(* IEC 61131-3 sources: 2026_Projet_YGO_ExcavatriceDragage/CODE/MAIN (part 2) *)

(* ---- PRG_09_Supervision.st ---- *)
(* ═══════════════════════════════════════════════════════════════
   🖥️ PRG_09_Supervision — Échanges IHM, Stubs et Initialisation Boot
   ───────────────────────────────────────────────────────────────
   ⚙️ Exécuté par la tâche PLC en position 9.
   ✅ Regroupe tout le mapping bidirectionnel GVL_IHM / GVL_PERSISTENT.
   ✅ Expose FaultMachineReset_IHM pour tous les programmes du domaine sécurité/métier.
   🔧 REX 2026-07-07 : séparation des resets — l'ancien MachineReset_IHM (unique, câblé sur
      TOUT y compris FB_Modes/FB_Cycle) est retiré. FaultMachineReset_IHM ne couvre plus que le
      domaine sécurité/métier (Winch, Safety, Encodeurs, Benne, Joystick, Translation) ;
      FB_Modes/FB_Cycle ont chacun leur propre Reset dédié (GVL_IHM.Modes.ModeReset côté
      PRG_04_Modes, CmdResetCycle_IHM côté PRG_05_Cycle) — jamais mélangés.
   ═══════════════════════════════════════════════════════════════ *)

PROGRAM PRG_09_Supervision
VAR_OUTPUT
    FaultMachineReset_IHM : BOOL; // 🔔 Acquittement défauts domaine sécurité/métier (OR des boutons HMI) — jamais Modes/Cycle
END_VAR
VAR
    instBlink1Hz : BLINK; // 🧩 Réutilisation lib Util (Partie3 §0) — horloge clignotement système
END_VAR

// === IMPLEMENTATION (corps du PROGRAM PRG_09_Supervision) ===

// ── 0. HORLOGE CLIGNOTEMENT SYSTÈME (GVL_Global.BlinkClock) ───────────────
// 🧩 Réutilisation lib Util (Partie3 §0) : bloc standard BLINK, pas de TON maison —
// gère nativement un rythme allumé/éteint ASYMÉTRIQUE (TimeHigh ≠ TimeLow), contrairement
// au motif TON manuel de FB_Output.st (symétrique 500/500, propre à l'option relais).
// 🔧 REX 2026-07-16 : durées réglables sans recompiler (GVL_PERSISTENT._BlinkTimeOn/_BlinkTimeOff,
// défaut 1s allumé / 800ms éteint) — un seul rythme partagé pour tous les voyants IHM/diag qui
// clignotent pareil.
// 💡 Un voyant a besoin d'un AUTRE rythme ? Instancier son propre BLINK localement (Util) avec
// ses propres TimeHigh/TimeLow — ne pas détourner ce bit partagé pour un rythme différent.
instBlink1Hz(
    ENABLE   := TRUE,
    TIMEHIGH := _BlinkTimeOn,
    TIMELOW  := _BlinkTimeOff
);
GVL_Global.BlinkClock := instBlink1Hz.OUT;

// ── 1. ACQUISITION DES DEMANDES / BOUTONS DE L'IHM ────────────────────────
GVL_Modes_Stub.ModeRequest_IHM         := GVL_IHM.Modes.ModeRequest;
GVL_Modes_Stub.SyncEnableRequest_IHM   := GVL_IHM.Sync.SyncEnableRequest; // 🔧 REX 2026-07-08 : renommé, polarité inversée
StubTranslationPositionSelect_IHM          := GVL_IHM.TranslationM3.SelectedTargetNum;

// Signal d'acquittement défauts domaine sécurité/métier — JAMAIS Modes/Cycle (REX 2026-07-07)
FaultMachineReset_IHM := GVL_IHM.Modes.FaultMachineReset
                    OR GVL_IHM.M1TreuilRetenue.CmdReset
                    OR GVL_IHM.M2TreuilBucket.CmdReset
                    OR GVL_IHM.Bucket.CmdReset;

// 🔴 REX 2026-07-07 : au moins un défaut actif dans le domaine couvert par FaultMachineReset_IHM
// (même périmètre exact que les 17 blocs alimentés par ce reset — voir bandeau en tête de fichier).
// Sert à savoir, côté IHM, quand un appui sur FaultMachineReset est utile/attendu.
GVL_IHM.Modes.AnyFaultActive :=
       PRG_01_Diagnostics.instDiagCanOpen.Error
    OR PRG_01_Diagnostics.instDiagEthercat.Error
    OR PRG_01_Diagnostics.FB_Joystick_0.Error
    OR (NOT PRG_04_Modes.instModes.InhibitM1 AND (
           PRG_02_Encoders.instEncoderAbsM1.Error
        OR PRG_02_Encoders.instHomingM1.Error
        OR PRG_02_Encoders.instEncoderSafetyM1.Error
        OR PRG_03_Safety.instSafetyWinchM1.Error
        OR PRG_06_WinchControl.instWinchM1.Error
    ))
    OR (NOT PRG_04_Modes.instModes.InhibitM2 AND (
           PRG_02_Encoders.instEncoderAbsM2.Error
        OR PRG_02_Encoders.instHomingM2.Error
        OR PRG_02_Encoders.instEncoderSafetyM2.Error
        OR PRG_03_Safety.instSafetyWinchM2.Error
        OR PRG_06_WinchControl.instWinchM2.Error
    ))
    OR PRG_03_Safety.instSafetyTranslationM3.Error
    OR PRG_06_WinchControl.instWinchSync.Error
    OR PRG_06_WinchControl.instBucket.Error
    OR PRG_07_TranslationControl.instTranslationM3.Error
    OR PRG_10_Outputs.RedundancyTestFailed
    OR PRG_10_Outputs.EmergencyArmingFailed;

// 🧨 REX 2026-07-07 : remontée IHM de la coupure puissance amont — polarité "alarme" (TRUE=
// problème), PAS celle de PowerCutOff_A_RQ (qui est en fail-safe maintenu, TRUE=OK depuis
// l'inversion de polarité). On relit directement les .PowerCutOff sources, pas la sortie physique.
GVL_IHM.Modes.PowerCutOffActive := PRG_03_Safety.instSafetyWinchM1.PowerCutOff
                                 OR PRG_03_Safety.instSafetyWinchM2.PowerCutOff
                                 OR PRG_03_Safety.instSafetyTranslationM3.PowerCutOff
                                 OR GVL_IHM.Modes.CmdEmergencyCutOff;

// 🆕 REX 2026-07-08 : thermique frein commun M1/M2/M3 — signal UNIQUE (1 seul fil, pas de sens à
// le dupliquer par axe), remonté une seule fois au niveau global GVL_IHM (même principe que
// TopPositionSensorActive ci-dessus, PAS dans WinchM1/WinchM2/Translation).
GVL_IHM.Commun.BrakeThermalFault := NOT PRG_00_Inputs.BrakeThermalFeedback;
GVL_IHM.Commun.PhaseRotationFault := NOT PRG_00_Inputs.PhaseRotationOk; // 🆕 REX 2026-07-08 — commun M1/M2/M3, invisible IHM avant

// 🔧 REX 2026-07-07 — Séquence réarmement AU (voir DOC/AF_Partie1 v1.5 §Sécurité électrique)
// EmergencyArmingBusy couvre TOUTE la séquence (auto-test A/B + pulse + confirmation + verrouillage),
// pas seulement le pulse — ArmingSeqStep<>0 englobe déjà tout sauf le verrouillage final.
GVL_IHM.Modes.EmergencyChainOk    := PRG_00_Inputs.EmergencyChain;
GVL_IHM.Modes.PowerContactorOk    := PRG_00_Inputs.EmergencyStopOk;
GVL_IHM.Modes.EmergencyArmingBusy := (PRG_10_Outputs.ArmingSeqStep <> 0) OR PRG_10_Outputs.EmergencyArmingLockoutActive;
GVL_IHM.Modes.EmergencyArmable    := PRG_00_Inputs.EmergencyChain
                                    AND (PRG_10_Outputs.ArmingSeqStep = 0)
                                    AND NOT PRG_10_Outputs.EmergencyArmingLockoutActive
                                    AND NOT PRG_10_Outputs.RedundancyTestFailed;
GVL_IHM.Modes.RedundancyTestFailed := PRG_10_Outputs.RedundancyTestFailed;
GVL_IHM.Modes.EmergencyArmingFailed := PRG_10_Outputs.EmergencyArmingFailed;

// 🔧 REX 2026-07-07 : ancien pont IF/ELSIF vers GVL_Encoder_Stub supprimé (bugué — ne pouvait
// homer qu'un seul treuil à la fois). GVL_IHM.M1TreuilRetenue/M2.CmdHome sont désormais câblés
// directement dans PRG_02_Encoders.st (instHomingM1/M2.Home) — homing simultané possible.

// ℹ️ Calibrate joystick : lu directement depuis GVL_IHM.JoystickJOY1.Calibrate dans PRG_01_Diagnostics (ligne 48)
// PRG_01_Diagnostics.FB_Joystick_0.Calibrate := GVL_IHM.JoystickJOY1.Calibrate;  // ❌ supprimé : VAR locale non accessible en écriture (C0037)

// ── 2. INITIALISATION IHM DEPUIS GVL_PERSISTENT (Boot) ───────────────────
IF GVL_IHM.M1TreuilRetenue.TopSensorPositionM = 0.0 THEN
    GVL_IHM.M1TreuilRetenue.TopSensorPositionM  := _HomingTargetM1_M;
    GVL_IHM.M1TreuilRetenue.MaxStepDescente     := _WinchMaxStepDescent; // 🔧 REX 2026-07-08 : commun M1/M2
    GVL_IHM.M1TreuilRetenue.RampAccelRate       := _WinchM1RampAccelRate_Pct;
    GVL_IHM.M1TreuilRetenue.RampDecelNormalRate := _WinchM1RampDecelNormal_Pct;
    GVL_IHM.M1TreuilRetenue.RampDecelFastRate   := _WinchM1RampDecelFast_Pct;
    GVL_IHM.M1TreuilRetenue.CableLimitDescentM  := _CableLimitM1Descent_M;
    GVL_IHM.M1TreuilRetenue.CableLimitAscentM   := _CableLimitM1Ascent_M; // 🆕 REX 2026-07-15 (6)
    GVL_IHM.M1TreuilRetenue.SlowdownDistanceM   := _WinchSlowdownDistance_M;
    GVL_IHM.M1TreuilRetenue.SlowSpeedPct        := _WinchSlowSpeed_Pct;
END_IF;

IF GVL_IHM.M2TreuilBucket.TopSensorPositionM = 0.0 THEN
    GVL_IHM.M2TreuilBucket.TopSensorPositionM  := _HomingTargetM2_M;
    GVL_IHM.M2TreuilBucket.MaxStepDescente     := _WinchMaxStepDescent; // 🔧 REX 2026-07-08 : commun M1/M2
    GVL_IHM.M2TreuilBucket.RampAccelRate       := _WinchM2RampAccelRate_Pct;
    GVL_IHM.M2TreuilBucket.RampDecelNormalRate := _WinchM2RampDecelNormal_Pct;
    GVL_IHM.M2TreuilBucket.RampDecelFastRate   := _WinchM2RampDecelFast_Pct;
    GVL_IHM.M2TreuilBucket.CableLimitDescentM  := _CableLimitM2Descent_M;
    GVL_IHM.M2TreuilBucket.CableLimitAscentM   := _CableLimitM2Ascent_M; // 🆕 REX 2026-07-15 (6)
    GVL_IHM.M2TreuilBucket.SlowdownDistanceM   := _WinchSlowdownDistance_M;
    GVL_IHM.M2TreuilBucket.SlowSpeedPct        := _WinchSlowSpeed_Pct;
END_IF;

IF GVL_IHM.Sync.SyncToleranceM = 0.0 THEN
    GVL_IHM.Sync.SyncToleranceM         := _WinchSyncTolerance_M;
END_IF;

IF GVL_IHM.Bucket.Config.OffsetOpenM = 0.0 AND GVL_IHM.Bucket.Config.OffsetCloseM = 0.0 THEN
    GVL_IHM.Bucket.Config := _BucketConfig;
    GVL_IHM.Bucket.TimeoutDuration := T#30s;
END_IF;

IF GVL_IHM.Commun.LimitLegalDepthMinAllowed = 0.0 THEN
    GVL_IHM.Commun.LimitLegalDepthMinAllowed := _LimitLegalDepthMinAllowed_M;
    GVL_IHM.Commun.LimitLegalEnabled         := _LimitLegalEnabled;
END_IF;

// 🆕 REX 2026-07-15 (10) — BUG CORRIGÉ (retour terrain) : WinchMaxStepFwd/Rev (essais progressifs
// IHM_MANU, TEMPORAIRE) n'avaient jamais de boot-init, contrairement à tous les autres réglages
// IHM ci-dessus — restaient à 0 (défaut INT) en permanence. Le bornage de PRG_06_WinchControl
// traitait ce 0 comme "invalide" et le remplaçait SILENCIEUSEMENT par 5 (aucune restriction),
// sans jamais corriger l'affichage IHM : l'opérateur voyait "0" (lu comme restrictif) alors que
// la vitesse réellement appliquée était pleine échelle — d'où les contacteurs qui commutaient
// normalement malgré un "0" à l'écran. GVL_IHM.IHM_MANU est déjà RETAIN (ST_IHM_MANU) — pas besoin
// de miroir GVL_PERSISTENT (dérogation temporaire, pas un réglage machine permanent, voir
// IHM_MANU_Journal_Modifications.md §10).
IF GVL_IHM.IHM_MANU.WinchMaxStepFwd = 0 THEN
    GVL_IHM.IHM_MANU.WinchMaxStepFwd := 5;
END_IF;
IF GVL_IHM.IHM_MANU.WinchMaxStepRev = 0 THEN
    GVL_IHM.IHM_MANU.WinchMaxStepRev := 2;
END_IF;

IF GVL_IHM.Modes.ModeRequest = E_Mode.DISABLE THEN
    GVL_IHM.Modes.ModeRequest := E_Mode.MAINT_N1;
END_IF;

// ── 3. PROPAGATION DES RÉGLAGES IHM → PERSISTANCE ───────────────────────
_HomingTargetM1_M           := GVL_IHM.M1TreuilRetenue.TopSensorPositionM;
_HomingTargetM2_M           := GVL_IHM.M2TreuilBucket.TopSensorPositionM;
// 🔧 REX 2026-07-08 : MaxStepDescente désormais commun M1/M2 — voir bloc miroir bidirectionnel
// ci-dessous (même pattern que CableLimitDescentM/SlowdownDistanceM/SlowSpeedPct), plus de
// propagation à sens unique séparée par treuil ici.
_WinchM1RampAccelRate_Pct   := GVL_IHM.M1TreuilRetenue.RampAccelRate;
_WinchM1RampDecelNormal_Pct := GVL_IHM.M1TreuilRetenue.RampDecelNormalRate;
_WinchM1RampDecelFast_Pct   := GVL_IHM.M1TreuilRetenue.RampDecelFastRate;
_WinchM2RampAccelRate_Pct   := GVL_IHM.M2TreuilBucket.RampAccelRate;
_WinchM2RampDecelNormal_Pct := GVL_IHM.M2TreuilBucket.RampDecelNormalRate;
_WinchM2RampDecelFast_Pct   := GVL_IHM.M2TreuilBucket.RampDecelFastRate;
// ⚠️ REX 2026-07-08 (5) — PIÈGE pont IHM→PERSISTENT découvert lors de l'audit : cette ligne
// écrase _WinchSyncTolerance_M avec GVL_IHM.Sync.SyncToleranceM À CHAQUE SCAN.
// Si on change UNIQUEMENT la valeur par défaut dans GVL_PERSISTENT.st (ou ST_SyncHMI.st), ça ne
// suffit pas : la valeur restaurée au boot (bloc §2 ci-dessus, `IF ... = 0.0 THEN`) ne s'applique
// que si le RETAIN IHM est à 0.0 (premier démarrage) — sinon l'ancienne valeur IHM re-propage ici
// et écrase silencieusement toute nouvelle valeur par défaut au scan suivant.
_WinchSyncTolerance_M       := GVL_IHM.Sync.SyncToleranceM;
_BucketConfig              := GVL_IHM.Bucket.Config;

// 🔧 REX 2026-07-08 (demande utilisateur) : MaxStepDescente commun M1/M2 — même profil de
// déplacement des 2 treuils, même pattern miroir que CableLimitDescentM ci-dessous.
IF GVL_IHM.M1TreuilRetenue.MaxStepDescente <> _WinchMaxStepDescent THEN
    _WinchMaxStepDescent := GVL_IHM.M1TreuilRetenue.MaxStepDescente;
ELSIF GVL_IHM.M2TreuilBucket.MaxStepDescente <> _WinchMaxStepDescent THEN
    _WinchMaxStepDescent := GVL_IHM.M2TreuilBucket.MaxStepDescente;
END_IF;
GVL_IHM.M1TreuilRetenue.MaxStepDescente := _WinchMaxStepDescent;
GVL_IHM.M2TreuilBucket.MaxStepDescente := _WinchMaxStepDescent;

IF GVL_IHM.M1TreuilRetenue.CableLimitDescentM <> _CableLimitM1Descent_M THEN
    _CableLimitM1Descent_M := GVL_IHM.M1TreuilRetenue.CableLimitDescentM;
END_IF;
GVL_IHM.M1TreuilRetenue.CableLimitDescentM := _CableLimitM1Descent_M;

IF GVL_IHM.M2TreuilBucket.CableLimitDescentM <> _CableLimitM2Descent_M THEN
    _CableLimitM2Descent_M := GVL_IHM.M2TreuilBucket.CableLimitDescentM;
END_IF;
GVL_IHM.M2TreuilBucket.CableLimitDescentM := _CableLimitM2Descent_M;

// 🆕 REX 2026-07-15 (6) — même pattern miroir bidirectionnel que CableLimitDescentM ci-dessus.
IF GVL_IHM.M1TreuilRetenue.CableLimitAscentM <> _CableLimitM1Ascent_M THEN
    _CableLimitM1Ascent_M := GVL_IHM.M1TreuilRetenue.CableLimitAscentM;
END_IF;
GVL_IHM.M1TreuilRetenue.CableLimitAscentM := _CableLimitM1Ascent_M;

IF GVL_IHM.M2TreuilBucket.CableLimitAscentM <> _CableLimitM2Ascent_M THEN
    _CableLimitM2Ascent_M := GVL_IHM.M2TreuilBucket.CableLimitAscentM;
END_IF;
GVL_IHM.M2TreuilBucket.CableLimitAscentM := _CableLimitM2Ascent_M;

IF GVL_IHM.M1TreuilRetenue.SlowdownDistanceM <> _WinchSlowdownDistance_M THEN
    _WinchSlowdownDistance_M := GVL_IHM.M1TreuilRetenue.SlowdownDistanceM;
ELSIF GVL_IHM.M2TreuilBucket.SlowdownDistanceM <> _WinchSlowdownDistance_M THEN
    _WinchSlowdownDistance_M := GVL_IHM.M2TreuilBucket.SlowdownDistanceM;
END_IF;
GVL_IHM.M1TreuilRetenue.SlowdownDistanceM := _WinchSlowdownDistance_M;
GVL_IHM.M2TreuilBucket.SlowdownDistanceM := _WinchSlowdownDistance_M;

IF GVL_IHM.M1TreuilRetenue.SlowSpeedPct <> _WinchSlowSpeed_Pct THEN
    _WinchSlowSpeed_Pct := GVL_IHM.M1TreuilRetenue.SlowSpeedPct;
ELSIF GVL_IHM.M2TreuilBucket.SlowSpeedPct <> _WinchSlowSpeed_Pct THEN
    _WinchSlowSpeed_Pct := GVL_IHM.M2TreuilBucket.SlowSpeedPct;
END_IF;
GVL_IHM.M1TreuilRetenue.SlowSpeedPct := _WinchSlowSpeed_Pct;
GVL_IHM.M2TreuilBucket.SlowSpeedPct := _WinchSlowSpeed_Pct;

_LimitLegalDepthMinAllowed_M := GVL_IHM.Commun.LimitLegalDepthMinAllowed;
_LimitLegalEnabled         := GVL_IHM.Commun.LimitLegalEnabled;
// 🔧 REX 2026-07-07 : plus de garde Mode=SEMI_AUTO, cohérent avec PRG_06_WinchControl.st §5
// (la limite légale s'applique désormais dans tous les modes dès qu'elle est activée).
GVL_IHM.Commun.LimitLegalReached         := _LimitLegalEnabled
                                            AND ((NOT PRG_04_Modes.instModes.InhibitM1 AND (PRG_02_Encoders.instEncoderScaleM1.CablePosM <= _LimitLegalDepthMinAllowed_M))
                                                 OR (NOT PRG_04_Modes.instModes.InhibitM2 AND (PRG_02_Encoders.instEncoderScaleM2.CablePosM <= _LimitLegalDepthMinAllowed_M)));

GVL_IHM.Commun.TopPositionSensorActive   := NOT PRG_00_Inputs.TopPositionSensor;

// ── 4. BYPASS DE SIMULATION POUR L'IHM (état effectif par device, voir AF_Partie13) ──────
GVL_IHM.M1TreuilRetenue.BypassContactorFeedback := GVL_Simulation.SimulationModeActive AND NOT GVL_Simulation.ContactorFeedbackM1_IsReal;
GVL_IHM.M2TreuilBucket.BypassContactorFeedback := GVL_Simulation.SimulationModeActive AND NOT GVL_Simulation.ContactorFeedbackM2_IsReal;
GVL_IHM.TranslationM3.BypassContactorFeedback := GVL_Simulation.SimulationModeActive AND NOT GVL_Simulation.ContactorFeedbackM3_IsReal;
GVL_IHM.M1TreuilRetenue.BypassSlackCable        := GVL_Simulation.SimulationModeActive AND NOT GVL_Simulation.SlackCableSwitch_IsReal;
GVL_IHM.M2TreuilBucket.BypassSlackCable        := GVL_Simulation.SimulationModeActive AND NOT GVL_Simulation.SlackCableSwitch_IsReal;
GVL_IHM.M1TreuilRetenue.BypassTopPositionSensor := GVL_Simulation.SimulationModeActive AND NOT GVL_Simulation.TopPositionSensor_IsReal;
GVL_IHM.M2TreuilBucket.BypassTopPositionSensor := GVL_Simulation.SimulationModeActive AND NOT GVL_Simulation.TopPositionSensor_IsReal;

// ── 5. MAPPING ÉTATS TREUIL M1 → IHM ─────────────────────────────────────
GVL_IHM.M1TreuilRetenue.PositionM                := PRG_02_Encoders.instEncoderScaleM1.CablePosM;
GVL_IHM.M1TreuilRetenue.SpeedRefPct              := PRG_06_WinchControl.instWinchM1.SpeedRamp.Current;
GVL_IHM.M1TreuilRetenue.StepNumber               := PRG_06_WinchControl.instWinchM1.StepNumber;
GVL_IHM.M1TreuilRetenue.FBState                  := PRG_06_WinchControl.instWinchM1.State;
GVL_IHM.M1TreuilRetenue.Ready                    := PRG_06_WinchControl.instWinchM1.Ready;
GVL_IHM.M1TreuilRetenue.Busy                     := PRG_06_WinchControl.instWinchM1.Busy;
GVL_IHM.M1TreuilRetenue.Done                     := PRG_06_WinchControl.instWinchM1.Done;
GVL_IHM.M1TreuilRetenue.Error                    := PRG_06_WinchControl.instWinchM1.Error;
GVL_IHM.M1TreuilRetenue.ErrorId                  := PRG_06_WinchControl.instWinchM1.ErrorId;
GVL_IHM.M1TreuilRetenue.RelayFwd                 := PRG_06_WinchControl.instWinchM1.RelayFwd;
GVL_IHM.M1TreuilRetenue.RelayRev                 := PRG_06_WinchControl.instWinchM1.RelayRev;
GVL_IHM.M1TreuilRetenue.Contactor1               := PRG_06_WinchControl.instWinchM1.Contactor1;
GVL_IHM.M1TreuilRetenue.Contactor2               := PRG_06_WinchControl.instWinchM1.Contactor2;
GVL_IHM.M1TreuilRetenue.Contactor3               := PRG_06_WinchControl.instWinchM1.Contactor3;
GVL_IHM.M1TreuilRetenue.Contactor4               := PRG_06_WinchControl.instWinchM1.Contactor4;
GVL_IHM.M1TreuilRetenue.BrakeCmd                 := PRG_06_WinchControl.instWinchM1.BrakeCmd;
GVL_IHM.M1TreuilRetenue.Homed                    := PRG_02_Encoders.instHomingM1.Homed;
GVL_IHM.M1TreuilRetenue.SafeStopActive           := PRG_03_Safety.instSafetyWinchM1.SafeStop;
GVL_IHM.M1TreuilRetenue.ForbidDescentActive      := PRG_06_WinchControl.ForbidDescentM1_Active;
GVL_IHM.M1TreuilRetenue.ForbidAscentActive       := PRG_03_Safety.instSafetyWinchM1.ForbidAscent;
GVL_IHM.M1TreuilRetenue.SlackCableDetected       := NOT PRG_00_Inputs.SlackCableSwitch;
GVL_IHM.M1TreuilRetenue.ThermalFault             := NOT PRG_00_Inputs.M1ThermalFeedback;
GVL_IHM.M1TreuilRetenue.EncoderFault             := NOT PRG_02_Encoders.instEncoderAbsM1.EncoderAvailable OR PRG_02_Encoders.instEncoderSafetyM1.EncoderIncoherent;
GVL_IHM.M1TreuilRetenue.CableLimitDescentReached := (PRG_03_Safety.instSafetyWinchM1.ErrorId AND 16#0040) <> 16#0000;
GVL_IHM.M1TreuilRetenue.CableLimitAscentReached  := PRG_06_WinchControl.CableLimitAscentM1Reached; // 🆕 REX 2026-07-15 (8)
GVL_IHM.M1TreuilRetenue.ContactorsCheck          := PRG_06_WinchControl.instWinchM1.ContactorsCheck; // 🔧 REX 2026-07-07
GVL_IHM.M1TreuilRetenue.BrakeContactorCheck      := PRG_06_WinchControl.instWinchM1.BrakeContactorCheck;

GVL_IHM.M1TreuilRetenue.Encoder.RawPos           := PRG_02_Encoders.instEncoderAbsM1.RawPos;
GVL_IHM.M1TreuilRetenue.Encoder.Alarms           := PRG_02_Encoders.instEncoderAbsM1.AlarmsIn;
GVL_IHM.M1TreuilRetenue.Encoder.Warnings         := PRG_02_Encoders.instEncoderAbsM1.WarningsIn;
GVL_IHM.M1TreuilRetenue.Encoder.SlaveOperational := PRG_02_Encoders.instEncoderAbsM1.SlaveOperational;
GVL_IHM.M1TreuilRetenue.Encoder.PresetTriggerCmd := PRG_02_Encoders.instEncoderAbsM1.PresetTriggerCmd;
GVL_IHM.M1TreuilRetenue.Encoder.PresetValueOut   := PRG_02_Encoders.instEncoderAbsM1.PresetValueOut;
GVL_IHM.M1TreuilRetenue.Encoder.Error            := PRG_02_Encoders.instEncoderAbsM1.Error;
GVL_IHM.M1TreuilRetenue.Encoder.ErrorId          := PRG_02_Encoders.instEncoderAbsM1.ErrorId;
GVL_IHM.M1TreuilRetenue.SafetyError              := PRG_03_Safety.instSafetyWinchM1.Error;
GVL_IHM.M1TreuilRetenue.SafetyErrorId            := PRG_03_Safety.instSafetyWinchM1.ErrorId;
GVL_IHM.M1TreuilRetenue.MecaADriftM              := PRG_03_Safety.instSafetyWinchM1.MecaADriftM;      // 🆕 REX 2026-07-08
GVL_IHM.M1TreuilRetenue.MecaCDriftM              := PRG_03_Safety.instSafetyWinchM1.MecaCDriftM;      // 🆕 REX 2026-07-08
GVL_IHM.M1TreuilRetenue.MecaBElapsedTime         := PRG_03_Safety.instSafetyWinchM1.MecaBElapsedTime; // 🆕 REX 2026-07-08
GVL_IHM.M1TreuilRetenue.InhibitActive            := PRG_04_Modes.instModes.InhibitM1; // 🆕 REX 2026-07-08

// ── 6. MAPPING ÉTATS TREUIL M2 → IHM ─────────────────────────────────────
GVL_IHM.M2TreuilBucket.PositionM                := PRG_02_Encoders.instEncoderScaleM2.CablePosM;
GVL_IHM.M2TreuilBucket.SpeedRefPct              := PRG_06_WinchControl.instWinchM2.SpeedRamp.Current;
GVL_IHM.M2TreuilBucket.StepNumber               := PRG_06_WinchControl.instWinchM2.StepNumber;
GVL_IHM.M2TreuilBucket.FBState                  := PRG_06_WinchControl.instWinchM2.State;
GVL_IHM.M2TreuilBucket.Ready                    := PRG_06_WinchControl.instWinchM2.Ready;
GVL_IHM.M2TreuilBucket.Busy                     := PRG_06_WinchControl.instWinchM2.Busy;
GVL_IHM.M2TreuilBucket.Done                     := PRG_06_WinchControl.instWinchM2.Done;
GVL_IHM.M2TreuilBucket.Error                    := PRG_06_WinchControl.instWinchM2.Error;
GVL_IHM.M2TreuilBucket.ErrorId                  := PRG_06_WinchControl.instWinchM2.ErrorId;
GVL_IHM.M2TreuilBucket.RelayFwd                 := PRG_06_WinchControl.instWinchM2.RelayFwd;
GVL_IHM.M2TreuilBucket.RelayRev                 := PRG_06_WinchControl.instWinchM2.RelayRev;
GVL_IHM.M2TreuilBucket.Contactor1               := PRG_06_WinchControl.instWinchM2.Contactor1;
GVL_IHM.M2TreuilBucket.Contactor2               := PRG_06_WinchControl.instWinchM2.Contactor2;
GVL_IHM.M2TreuilBucket.Contactor3               := PRG_06_WinchControl.instWinchM2.Contactor3;
GVL_IHM.M2TreuilBucket.Contactor4               := PRG_06_WinchControl.instWinchM2.Contactor4;
GVL_IHM.M2TreuilBucket.BrakeCmd                 := PRG_06_WinchControl.instWinchM2.BrakeCmd;
GVL_IHM.M2TreuilBucket.Homed                    := PRG_02_Encoders.instHomingM2.Homed;
GVL_IHM.M2TreuilBucket.SafeStopActive           := PRG_03_Safety.instSafetyWinchM2.SafeStop;
GVL_IHM.M2TreuilBucket.ForbidDescentActive      := PRG_06_WinchControl.ForbidDescentM2_Active;
GVL_IHM.M2TreuilBucket.ForbidAscentActive       := PRG_03_Safety.instSafetyWinchM2.ForbidAscent;
GVL_IHM.M2TreuilBucket.SlackCableDetected       := NOT PRG_00_Inputs.SlackCableSwitch;
GVL_IHM.M2TreuilBucket.ThermalFault             := NOT PRG_00_Inputs.M2ThermalFeedback;
GVL_IHM.M2TreuilBucket.EncoderFault             := NOT PRG_02_Encoders.instEncoderAbsM2.EncoderAvailable OR PRG_02_Encoders.instEncoderSafetyM2.EncoderIncoherent;
GVL_IHM.M2TreuilBucket.CableLimitDescentReached := (PRG_03_Safety.instSafetyWinchM2.ErrorId AND 16#0040) <> 16#0000;
GVL_IHM.M2TreuilBucket.CableLimitAscentReached  := PRG_06_WinchControl.CableLimitAscentM2Reached; // 🆕 REX 2026-07-15 (8)
GVL_IHM.M2TreuilBucket.ContactorsCheck          := PRG_06_WinchControl.instWinchM2.ContactorsCheck; // 🔧 REX 2026-07-07
GVL_IHM.M2TreuilBucket.BrakeContactorCheck      := PRG_06_WinchControl.instWinchM2.BrakeContactorCheck;

GVL_IHM.M2TreuilBucket.Encoder.RawPos           := PRG_02_Encoders.instEncoderAbsM2.RawPos;
GVL_IHM.M2TreuilBucket.Encoder.Alarms           := PRG_02_Encoders.instEncoderAbsM2.AlarmsIn;
GVL_IHM.M2TreuilBucket.Encoder.Warnings         := PRG_02_Encoders.instEncoderAbsM2.WarningsIn;
GVL_IHM.M2TreuilBucket.Encoder.SlaveOperational := PRG_02_Encoders.instEncoderAbsM2.SlaveOperational;
GVL_IHM.M2TreuilBucket.Encoder.PresetTriggerCmd := PRG_02_Encoders.instEncoderAbsM2.PresetTriggerCmd;
GVL_IHM.M2TreuilBucket.Encoder.PresetValueOut   := PRG_02_Encoders.instEncoderAbsM2.PresetValueOut;
GVL_IHM.M2TreuilBucket.Encoder.Error            := PRG_02_Encoders.instEncoderAbsM2.Error;
GVL_IHM.M2TreuilBucket.Encoder.ErrorId          := PRG_02_Encoders.instEncoderAbsM2.ErrorId;
GVL_IHM.M2TreuilBucket.SafetyError              := PRG_03_Safety.instSafetyWinchM2.Error;
GVL_IHM.M2TreuilBucket.SafetyErrorId            := PRG_03_Safety.instSafetyWinchM2.ErrorId;
GVL_IHM.M2TreuilBucket.MecaADriftM              := PRG_03_Safety.instSafetyWinchM2.MecaADriftM;      // 🆕 REX 2026-07-08
GVL_IHM.M2TreuilBucket.MecaCDriftM              := PRG_03_Safety.instSafetyWinchM2.MecaCDriftM;      // 🆕 REX 2026-07-08
GVL_IHM.M2TreuilBucket.MecaBElapsedTime         := PRG_03_Safety.instSafetyWinchM2.MecaBElapsedTime; // 🆕 REX 2026-07-08
GVL_IHM.M2TreuilBucket.InhibitActive            := PRG_04_Modes.instModes.InhibitM2; // 🆕 REX 2026-07-08

// ── 7. MAPPING ÉTATS BENNE → IHM ───────────────────────────────────────
GVL_IHM.Bucket.FBState          := PRG_06_WinchControl.instBucket.State;
GVL_IHM.Bucket.ActiveOffsetM    := PRG_06_WinchControl.instBucket.ActiveOffsetM;
GVL_IHM.Bucket.M2StartStop      := PRG_06_WinchControl.instBucket.M2_StartStop;
GVL_IHM.Bucket.M2Direction      := PRG_06_WinchControl.instBucket.M2_Direction;
GVL_IHM.Bucket.M2ForceSlowSpeed := PRG_06_WinchControl.instBucket.M2_ForceSlowSpeed;
GVL_IHM.Bucket.Ready            := PRG_06_WinchControl.instBucket.Ready;
GVL_IHM.Bucket.Busy             := PRG_06_WinchControl.instBucket.Busy;
GVL_IHM.Bucket.Done             := PRG_06_WinchControl.instBucket.Done;
GVL_IHM.Bucket.Error            := PRG_06_WinchControl.instBucket.Error;
GVL_IHM.Bucket.ErrorId          := PRG_06_WinchControl.instBucket.ErrorId;
GVL_IHM.Bucket.RemainingTravelM := PRG_06_WinchControl.instBucket.RemainingTravelM; // 🔧 REX 2026-07-07
GVL_IHM.Bucket.CloseReq         := PRG_06_WinchControl.instBucket.CloseReq; // 🆕 REX 2026-07-08
GVL_IHM.Bucket.OpenReq          := PRG_06_WinchControl.instBucket.OpenReq;  // 🆕 REX 2026-07-08
// 📊 REX 2026-07-07 : position M2 corrigée de l'offset actif — affichage bargraphe uniquement,
// doit être égale à GVL_IHM.M1TreuilRetenue.PositionM quand tout est nominal (voir bandeau ST_BucketHMI).
GVL_IHM.Bucket.M2PositionCorrected := PRG_02_Encoders.instEncoderScaleM2.CablePosM - PRG_06_WinchControl.instBucket.ActiveOffsetM;
GVL_IHM.Bucket.State            := _BucketState;

// ── 8. MAPPING ÉTATS SYNCHRONISATION → IHM ─────────────────────────────────
GVL_IHM.Sync.DeltaPosM  := PRG_06_WinchControl.instWinchSync.DeltaPosM;
GVL_IHM.Sync.SyncActive := PRG_06_WinchControl.instWinchSync.SyncActive;
GVL_IHM.Sync.SyncWarn   := PRG_06_WinchControl.instWinchSync.SyncWarn;
GVL_IHM.Sync.Ready      := PRG_06_WinchControl.instWinchSync.Ready;
GVL_IHM.Sync.Error      := PRG_06_WinchControl.instWinchSync.Error;
GVL_IHM.Sync.ErrorId    := PRG_06_WinchControl.instWinchSync.ErrorId;
GVL_IHM.Sync.State      := PRG_06_WinchControl.instWinchSync.State;

// ── 9. MAPPING ÉTATS TRANSLATION M3 → IHM ────────────────────────────────────
GVL_IHM.TranslationM3.FBState              := PRG_07_TranslationControl.instTranslationM3.State;
GVL_IHM.TranslationM3.Ready                := PRG_07_TranslationControl.instTranslationM3.Ready;
GVL_IHM.TranslationM3.Busy                 := PRG_07_TranslationControl.instTranslationM3.Busy;
GVL_IHM.TranslationM3.Done                 := PRG_07_TranslationControl.instTranslationM3.Done;
GVL_IHM.TranslationM3.Error                := PRG_07_TranslationControl.instTranslationM3.Error;
GVL_IHM.TranslationM3.ErrorId              := PRG_07_TranslationControl.instTranslationM3.ErrorId;
GVL_IHM.TranslationM3.BrakeCmd             := PRG_07_TranslationControl.instTranslationM3.BrakeCmd;
GVL_IHM.TranslationM3.BrakeFeedback        := PRG_00_Inputs.M3BrakeFeedback;
GVL_IHM.TranslationM3.PositionSensorTarget := PRG_07_TranslationControl.M3_PositionSensorTarget;
// 🔧 Diag variateur décodé (pas de bit-masking côté IHM) — StatusWord bit7=CommReady, bit0=PowerReady
GVL_IHM.TranslationM3.DriveCommReady       := PRG_00_Inputs.M3_StatusWord_Filtered.7 OR GVL_Simulation.SimulationModeActive;
GVL_IHM.TranslationM3.DrivePowerReady      := PRG_00_Inputs.M3_StatusWord_Filtered.0 OR GVL_Simulation.SimulationModeActive;
// 🔧 Source unique (PRG_00_Inputs), valable Auto ET Manu — remplace l'ex-doublon IHM_MANU.M3_FreqActual
GVL_IHM.TranslationM3.DriveActualFreqHz    := UINT_TO_REAL(PRG_00_Inputs.M3_ActualFrequencyHz_Filtered) / 100.0;
GVL_IHM.TranslationM3.SafetyError          := PRG_03_Safety.instSafetyTranslationM3.Error;
GVL_IHM.TranslationM3.SafetyErrorId        := PRG_03_Safety.instSafetyTranslationM3.ErrorId;
GVL_IHM.TranslationM3.SafetyErrorJoystick     := PRG_03_Safety.instSafetyTranslationM3.ErrorJoystick;
GVL_IHM.TranslationM3.SafetyErrorDriveComm    := PRG_03_Safety.instSafetyTranslationM3.ErrorDriveComm;
GVL_IHM.TranslationM3.SafetyErrorPhaseRotation:= PRG_03_Safety.instSafetyTranslationM3.ErrorPhaseRotation;
GVL_IHM.TranslationM3.SafetyErrorBrakeThermal := PRG_03_Safety.instSafetyTranslationM3.ErrorBrakeThermal;
GVL_IHM.TranslationM3.SafetyErrorMecaB        := PRG_03_Safety.instSafetyTranslationM3.ErrorMecaB;
GVL_IHM.TranslationM3.SafetyErrorMecaA        := PRG_03_Safety.instSafetyTranslationM3.ErrorMecaA;
GVL_IHM.TranslationM3.SafetyErrorLimitSwitch  := PRG_03_Safety.instSafetyTranslationM3.ErrorLimitSwitch;

// ── 10. MAPPING ÉTATS JOYSTICK → IHM ─────────────────────────────────────
GVL_IHM.JoystickJOY1.RawX       := JoyXRaw_ANA1;
GVL_IHM.JoystickJOY1.RawY       := JoyYRaw_ANA2;
GVL_IHM.JoystickJOY1.RawButton  := JoyBtnRaw;
GVL_IHM.JoystickJOY1.CmdX       := PRG_01_Diagnostics.FB_Joystick_0.AxisCmdX;
GVL_IHM.JoystickJOY1.CmdY       := PRG_01_Diagnostics.FB_Joystick_0.AxisCmdY;
GVL_IHM.JoystickJOY1.Online     := PRG_01_Diagnostics.instDiagCanOpen.DeviceJoystick.Online;
GVL_IHM.JoystickJOY1.Operational := PRG_01_Diagnostics.instDiagCanOpen.DeviceJoystick.Operational;
GVL_IHM.JoystickJOY1.Error       := PRG_01_Diagnostics.FB_Joystick_0.Error;
GVL_IHM.JoystickJOY1.ErrorId     := PRG_01_Diagnostics.FB_Joystick_0.ErrorId;

// ── 11. MAPPING SYSTEM / MODE → IHM ──────────────────────────────────────
GVL_IHM.Modes.CurrentMode     := PRG_04_Modes.instModes.Mode;
GVL_IHM.Modes.EmergencyStopOk := PRG_00_Inputs.EmergencyStopOk;

// ── 12. MAPPING DIAGNOSTICS BUS → IHM ────────────────────────────────────
GVL_IHM.Network.BusCanOpen  := PRG_01_Diagnostics.instDiagCanOpen.DeviceCanOpenMaster;
GVL_IHM.Network.Joystick    := PRG_01_Diagnostics.instDiagCanOpen.DeviceJoystick;
GVL_IHM.Network.CanError    := PRG_01_Diagnostics.instDiagCanOpen.Error;
GVL_IHM.Network.CanErrorId  := PRG_01_Diagnostics.instDiagCanOpen.ErrorId;

GVL_IHM.Network.BusEthercat := PRG_01_Diagnostics.instDiagEthercat.DeviceEthercatMaster;
GVL_IHM.Network.EncoderM1   := PRG_01_Diagnostics.instDiagEthercat.DeviceEncoderM1;
GVL_IHM.Network.EncoderM2   := PRG_01_Diagnostics.instDiagEthercat.DeviceEncoderM2;
GVL_IHM.Network.VariateurM3 := PRG_01_Diagnostics.instDiagEthercat.DeviceVariateur;
GVL_IHM.Network.EcatError   := PRG_01_Diagnostics.instDiagEthercat.Error;
GVL_IHM.Network.EcatErrorId := PRG_01_Diagnostics.instDiagEthercat.ErrorId;

(* ---- PRG_10_Outputs.st ---- *)
(* ═══════════════════════════════════════════════════════════════
   📤 PRG_10_Outputs — Écriture des SORTIES physiques (PROGRAMME)
   ───────────────────────────────────────────────────────────────
   📄 Doc : DOC/AF_Partie6_IO_Conditioning_v1.2.md §5
   ⚙️ Exécuté par la tâche PLC en position 10.
   ✅ Reçoit ses commandes en VAR_INPUT (écrites par le reste du code).
   ═══════════════════════════════════════════════════════════════ *)

PROGRAM PRG_10_Outputs
VAR_INPUT
    // ── 🪝 TREUIL M1 ─────────────────────────────────────────────────────────────────────
    M1RelayFwd        : BOOL;  // ⬆️ Relais MONTÉE M1 (NO) : TRUE=bobine ON, moteur monte | FALSE=arrêt ✅
    M1RelayRev        : BOOL;  // ⬇️ Relais DESCENTE M1 (NO) : TRUE=bobine ON, moteur descend | FALSE=arrêt ✅
    M1SpeedContactor1 : BOOL;  // 🐢 Contacteur vitesse 1 M1 — palier 1 lent (résistance max)
    M1SpeedContactor2 : BOOL;  // 🐇 Contacteur vitesse 2 M1 — palier 2
    M1SpeedContactor3 : BOOL;  // 🐇🐇 Contacteur vitesse 3 M1 — palier 3
    M1SpeedContactor4 : BOOL;  // 🚀 Contacteur vitesse 4 M1 — palier 4 pleine puissance
    M1BrakeCmd        : BOOL;  // 🔓 Frein M1 ⚠️INVERSÉ : TRUE=desserré/mouvement | FALSE=SERRÉ sécurité ✅

    // ── 🪝 TREUIL M2 (même logique que M1) ──────────────────────────────────────────────
    M2RelayFwd        : BOOL;  // ⬆️ Relais MONTÉE M2 (NO) : TRUE=bobine ON, moteur monte | FALSE=arrêt ✅
    M2RelayRev        : BOOL;  // ⬇️ Relais DESCENTE M2 (NO) : TRUE=bobine ON, moteur descend | FALSE=arrêt ✅
    M2SpeedContactor1 : BOOL;  // 🐢 Contacteur vitesse 1 M2 — palier 1 lent
    M2SpeedContactor2 : BOOL;  // 🐇 Contacteur vitesse 2 M2 — palier 2
    M2SpeedContactor3 : BOOL;  // 🐇🐇 Contacteur vitesse 3 M2 — palier 3
    M2SpeedContactor4 : BOOL;  // 🚀 Contacteur vitesse 4 M2 — palier 4 pleine puissance
    M2BrakeCmd        : BOOL;  // 🔓 Frein M2 ⚠️INVERSÉ : TRUE=desserré/mouvement | FALSE=SERRÉ sécurité ✅

    // ── ↔️ TRANSLATION M3 (sens/vitesse via variateur EtherCAT, TOR=frein uniquement) ────────
    TranslationBrakeCmd   : BOOL;  // 🔓 Frein M3 ⚠️INVERSÉ : TRUE=desserré/mouvement | FALSE=SERRÉ sécurité ✅
END_VAR
VAR_OUTPUT
    // 🔧 REX 2026-07-07 — état séquence réarmement AU, exposé pour affichage IHM (PRG_09_Supervision)
    EmergencyArmingPulseActive   : BOOL; // Pulse 1s en cours
    EmergencyArmingLockoutActive: BOOL; // Verrouillage 5s après pulse (mécanisme à ressort)
    ArmingSeqStep                : INT;  // 0=IDLE,1=TestA,2=RestoreA,3=TestB,4=RestoreB,5=Pulse,6=Confirm
    RedundancyTestFailed         : BOOL; // Canal A ou B non fonctionnel détecté à l'auto-test — bloque le réarmement
    EmergencyArmingFailed        : BOOL; // Impulsion envoyée mais contacteur puissance jamais confirmé
END_VAR
VAR
    // Instances de sortie
    instM1RelayFwd        : FB_Output;
    instM1RelayRev        : FB_Output;
    instM1SpeedContactor1 : FB_Output;
    instM1SpeedContactor2 : FB_Output;
    instM1SpeedContactor3 : FB_Output;
    instM1SpeedContactor4 : FB_Output;
    instM1BrakeCmd        : FB_Output;

    instM2RelayFwd        : FB_Output;
    instM2RelayRev        : FB_Output;
    instM2SpeedContactor1 : FB_Output;
    instM2SpeedContactor2 : FB_Output;
    instM2SpeedContactor3 : FB_Output;
    instM2SpeedContactor4 : FB_Output;
    instM2BrakeCmd        : FB_Output;

    instTranslationBrakeCmd   : FB_Output;
    instSafetyEmergencyManagement  : FB_Safety_EmergencyManagement;
    PowerCutOffReq            : BOOL;

    // ─────────  Début modification IHM_MANU  ─────────
    // 🆕 REX 2026-07-09 — Mode IHM_MANU (mise en service urgence, override direct sorties)
    ManuActive            : BOOL; // NOT GVL_IHM.IHM_MANU.ModeDisable (logique inversée, voir ST_IHM_MANU)
    // Détection de fronts montants pour priorité temporelle (Boutons HMI uniquement)
    TrigM1Fwd             : BOOL;
    TrigM1Rev             : BOOL;
    TrigM2Fwd             : BOOL;
    TrigM2Rev             : BOOL;
    TrigCoupledFwd        : BOOL;
    TrigCoupledRev        : BOOL;
    TrigM3Fwd             : BOOL;
    TrigM3Rev             : BOOL;
    // États au scan précédent (Boutons HMI uniquement)
    LastM1Fwd             : BOOL;
    LastM1Rev             : BOOL;
    LastM2Fwd             : BOOL;
    LastM2Rev             : BOOL;
    LastCoupledFwd        : BOOL;
    LastCoupledRev        : BOOL;
    LastM3Fwd             : BOOL;
    LastM3Rev             : BOOL;

    // Commandes brutes demandées (après aiguillage HMI / Joystick)
    M1Fwd_Demand          : BOOL;
    M1Rev_Demand          : BOOL;
    M2Fwd_Demand          : BOOL;
    M2Rev_Demand          : BOOL;
    CoupledFwd_Demand     : BOOL;
    CoupledRev_Demand     : BOOL;
    M3Fwd_Demand          : BOOL;
    M3Rev_Demand          : BOOL;

    // 🔧 REX 2026-07-15 (2) : rampe HMI locale (CycleTimeCalc/instHmiSpeedRamp/SpeedRefPct) et
    // décodage paliers (instManuSpeedStep/ActiveMaxStepFwd/Rev) RETIRÉS avec M1Fwd_Eff ci-dessus.
    // 🔧 REX 2026-07-16 : ex-M3Fwd_Eff/M3Rev_Eff/M3_ActiveFreqCmd/M3_DriveIsReal RETIRÉS — M3
    // piloté désormais par FB_Translation (PRG_07_TranslationControl §1bis), même principe que
    // M1/M2 (REX 2026-07-15 (2) ci-dessus) : plus besoin d'états effectifs locaux pour le bypass
    // M3_CommandWord (supprimé, voir fin de fichier).
    WinchMoving           : BOOL;         // 🚨 Au moins une commande de treuil HMI active (verrouillage aiguillage)
    M1_IsReal             : BOOL;         // ⚡ Indique si le treuil M1 est configuré comme réel
    M2_IsReal             : BOOL;         // ⚡ Indique si le treuil M2 est configuré comme réel
    M3_IsReal             : BOOL;         // ⚡ Indique si le translation M3 est configuré comme réel
    PowerCutOffActive_Eff : BOOL;         // ⚡ Indique si une coupure de puissance est active sur un équipement réel
    StartupNeutralOk      : BOOL := FALSE; // 🔒 Sécurité démarrage : exige le retour au neutre initial
    // ─────────  Fin modification IHM_MANU  ─────────
END_VAR

// === IMPLEMENTATION (corps du PROGRAM PRG_10_Outputs) ===

// ─────────  Début modification IHM_MANU  ─────────
// ═══════════════════════════════════════════════════════════════════════════
// 🚨 MODE IHM_MANU — override direct des sorties (mise en service urgence)
// ───────────────────────────────────────────────────────────────────────────
// 🆕 REX 2026-07-09 : logique inversée VOLONTAIRE — GVL_IHM.IHM_MANU.ModeDisable
// est non-RETAIN, donc FALSE à CHAQUE démarrage/download automate = mode Manu
// ACTIF d'origine, sans action opérateur. Il faut explicitement passer
// ModeDisable=TRUE pour rendre la main au programme fonctionnel normal
// (PRG_06_WinchControl/PRG_07_TranslationControl/PRG_03_Safety, intouchés).
// ⚠️ Aucune sécurité logicielle métier active en Manu (safety M1/M2/M3, synchro,
// limites logicielles, homing) — seuls les interlocks Fwd/Rev, K1-K4 ci-dessous,
// les fins de course benne, et la chaîne AU/PowerCutOff (§ plus bas, TOUJOURS
// active, non bypassée), protègent la machine et les personnes.
// 📍 Placé en tête de PRG_10_Outputs (position tâche 10, la plus en aval) : écrase
// les VAR_INPUT juste avant leur écriture réelle, APRÈS que PRG_06/07 (positions
// 6/7) les aient déjà remplis — le programme normal tourne dans le vide, ignoré.
ManuActive := NOT GVL_IHM.IHM_MANU.ModeDisable;

// Affichage position — utile même hors Manu pour vérifier le câblage codeur en direct
GVL_IHM.IHM_MANU.PositionM_M1 := PRG_02_Encoders.instEncoderScaleM1.CablePosM;
GVL_IHM.IHM_MANU.PositionM_M2 := PRG_02_Encoders.instEncoderScaleM2.CablePosM;

// 📊 Calcul de l'écart benne et des états de fin de course (delta = M1 - M2)
GVL_IHM.IHM_MANU.FdcBucketOpenEnable := GVL_IHM.IHM_MANU.FdcBucketOpen;
GVL_IHM.IHM_MANU.FdcBucketCloseEnable := GVL_IHM.IHM_MANU.FdcBucketClose;
GVL_IHM.IHM_MANU.BenneDelta := GVL_IHM.IHM_MANU.PositionM_M1 - GVL_IHM.IHM_MANU.PositionM_M2;
GVL_IHM.IHM_MANU.FdcBucketOpenActive  := GVL_IHM.IHM_MANU.FdcBucketOpenEnable AND (GVL_IHM.IHM_MANU.BenneDelta >= 0.0);
GVL_IHM.IHM_MANU.FdcBucketCloseActive := GVL_IHM.IHM_MANU.FdcBucketCloseEnable AND (GVL_IHM.IHM_MANU.BenneDelta <= -10.0);

IF ManuActive THEN
    // 1️⃣ Détection des nouveaux appuis sur boutons HMI (uniquement pour interlocks HMI)
    TrigM1Fwd      := GVL_IHM.IHM_MANU.M1_RelayFwd AND NOT LastM1Fwd;
    TrigM1Rev      := GVL_IHM.IHM_MANU.M1_RelayRev AND NOT LastM1Rev;
    TrigM2Fwd      := GVL_IHM.IHM_MANU.M2_RelayFwd AND NOT LastM2Fwd;
    TrigM2Rev      := GVL_IHM.IHM_MANU.M2_RelayRev AND NOT LastM2Rev;
    TrigCoupledFwd := GVL_IHM.IHM_MANU.M1_M2_RelayFwd AND NOT LastCoupledFwd;
    TrigCoupledRev := GVL_IHM.IHM_MANU.M1_M2_RelayRev AND NOT LastCoupledRev;
    TrigM3Fwd      := GVL_IHM.TranslationM3.ReqFwd AND NOT LastM3Fwd;
    TrigM3Rev      := GVL_IHM.TranslationM3.ReqRev AND NOT LastM3Rev;

    // 2️⃣ Interlocks de sécurité sur boutons HMI (Montée vs Descente)
    IF GVL_IHM.IHM_MANU.M1_RelayFwd AND GVL_IHM.IHM_MANU.M1_RelayRev THEN
        IF TrigM1Rev THEN
            GVL_IHM.IHM_MANU.M1_RelayRev := FALSE; (* Rejet Rev *)
        ELSIF TrigM1Fwd THEN
            GVL_IHM.IHM_MANU.M1_RelayFwd := FALSE; (* Rejet Fwd *)
        ELSE
            GVL_IHM.IHM_MANU.M1_RelayFwd := FALSE;
            GVL_IHM.IHM_MANU.M1_RelayRev := FALSE;
        END_IF;
    END_IF;

    IF GVL_IHM.IHM_MANU.M2_RelayFwd AND GVL_IHM.IHM_MANU.M2_RelayRev THEN
        IF TrigM2Rev THEN
            GVL_IHM.IHM_MANU.M2_RelayRev := FALSE;
        ELSIF TrigM2Fwd THEN
            GVL_IHM.IHM_MANU.M2_RelayFwd := FALSE;
        ELSE
            GVL_IHM.IHM_MANU.M2_RelayFwd := FALSE;
            GVL_IHM.IHM_MANU.M2_RelayRev := FALSE;
        END_IF;
    END_IF;

    IF GVL_IHM.IHM_MANU.M1_M2_RelayFwd AND GVL_IHM.IHM_MANU.M1_M2_RelayRev THEN
        IF TrigCoupledRev THEN
            GVL_IHM.IHM_MANU.M1_M2_RelayRev := FALSE;
        ELSIF TrigCoupledFwd THEN
            GVL_IHM.IHM_MANU.M1_M2_RelayFwd := FALSE;
        ELSE
            GVL_IHM.IHM_MANU.M1_M2_RelayFwd := FALSE;
            GVL_IHM.IHM_MANU.M1_M2_RelayRev := FALSE;
        END_IF;
    END_IF;

    IF GVL_IHM.TranslationM3.ReqFwd AND GVL_IHM.TranslationM3.ReqRev THEN
        IF TrigM3Rev THEN
            GVL_IHM.TranslationM3.ReqRev := FALSE;
        ELSIF TrigM3Fwd THEN
            GVL_IHM.TranslationM3.ReqFwd := FALSE;
        ELSE
            GVL_IHM.TranslationM3.ReqFwd := FALSE;
            GVL_IHM.TranslationM3.ReqRev := FALSE;
        END_IF;
    END_IF;

    // 3️⃣ Conflits boutons HMI entre mouvements Individuels et Couplés
    IF GVL_IHM.IHM_MANU.M1_M2_RelayFwd THEN
        IF GVL_IHM.IHM_MANU.M1_RelayRev THEN GVL_IHM.IHM_MANU.M1_RelayRev := FALSE; END_IF;
        IF GVL_IHM.IHM_MANU.M2_RelayRev THEN GVL_IHM.IHM_MANU.M2_RelayRev := FALSE; END_IF;
    END_IF;

    IF GVL_IHM.IHM_MANU.M1_M2_RelayRev THEN
        IF GVL_IHM.IHM_MANU.M1_RelayFwd THEN GVL_IHM.IHM_MANU.M1_RelayFwd := FALSE; END_IF;
        IF GVL_IHM.IHM_MANU.M2_RelayFwd THEN GVL_IHM.IHM_MANU.M2_RelayFwd := FALSE; END_IF;
    END_IF;

    IF (GVL_IHM.IHM_MANU.M1_RelayRev OR GVL_IHM.IHM_MANU.M2_RelayRev) AND GVL_IHM.IHM_MANU.M1_M2_RelayFwd THEN
        GVL_IHM.IHM_MANU.M1_M2_RelayFwd := FALSE;
    END_IF;

    IF (GVL_IHM.IHM_MANU.M1_RelayFwd OR GVL_IHM.IHM_MANU.M2_RelayFwd) AND GVL_IHM.IHM_MANU.M1_M2_RelayRev THEN
        GVL_IHM.IHM_MANU.M1_M2_RelayRev := FALSE;
    END_IF;

    // 4️⃣ Aiguillage de la commande de mouvement (HMI vs Joystick CANopen)
    M1_IsReal := NOT GVL_Simulation.SimulationModeActive OR GVL_Simulation.EncoderM1_IsReal OR GVL_Simulation.ContactorFeedbackM1_IsReal OR GVL_Simulation.ThermalM1_IsReal;
    M2_IsReal := NOT GVL_Simulation.SimulationModeActive OR GVL_Simulation.EncoderM2_IsReal OR GVL_Simulation.ContactorFeedbackM2_IsReal OR GVL_Simulation.ThermalM2_IsReal;
    M3_IsReal := NOT GVL_Simulation.SimulationModeActive OR GVL_Simulation.VariateurM3_IsReal OR GVL_Simulation.ContactorFeedbackM3_IsReal OR GVL_Simulation.TranslationPosition_IsReal;
    PowerCutOffActive_Eff := (M1_IsReal AND PRG_03_Safety.instSafetyWinchM1.PowerCutOff)
                             OR (M2_IsReal AND PRG_03_Safety.instSafetyWinchM2.PowerCutOff)
                             OR (M3_IsReal AND PRG_03_Safety.instSafetyTranslationM3.PowerCutOff);
    // ⚡ Clamp de sécurité sur la consigne saisie par l'opérateur (limité par le plafond absolu persistant)
    IF GVL_IHM.TranslationM3.FreqSetpointHz > _TranslationMaxFreq_Hz THEN
        GVL_IHM.TranslationM3.FreqSetpointHz := _TranslationMaxFreq_Hz;
    ELSIF GVL_IHM.TranslationM3.FreqSetpointHz < 0.0 THEN
        GVL_IHM.TranslationM3.FreqSetpointHz := 0.0;
    END_IF;

    IF GVL_IHM.IHM_MANU.JoystickSelect THEN
        // Commandes via le Joystick CANopen (arbitrées selon le mode de sécurité de FB_Modes, cf. TASK-0001)
        M1Fwd_Demand := (PRG_04_Modes.instModes.JoystickWinchSelectArbitrated = 1) AND (PRG_01_Diagnostics.FB_Joystick_0.AxisCmdY.Direction = 1);
        M1Rev_Demand := (PRG_04_Modes.instModes.JoystickWinchSelectArbitrated = 1) AND (PRG_01_Diagnostics.FB_Joystick_0.AxisCmdY.Direction = -1);

        M2Fwd_Demand := (PRG_04_Modes.instModes.JoystickWinchSelectArbitrated = 2) AND (PRG_01_Diagnostics.FB_Joystick_0.AxisCmdY.Direction = 1);
        M2Rev_Demand := (PRG_04_Modes.instModes.JoystickWinchSelectArbitrated = 2) AND (PRG_01_Diagnostics.FB_Joystick_0.AxisCmdY.Direction = -1);

        CoupledFwd_Demand := (PRG_04_Modes.instModes.JoystickWinchSelectArbitrated = 3) AND (PRG_01_Diagnostics.FB_Joystick_0.AxisCmdY.Direction = 1);
        CoupledRev_Demand := (PRG_04_Modes.instModes.JoystickWinchSelectArbitrated = 3) AND (PRG_01_Diagnostics.FB_Joystick_0.AxisCmdY.Direction = -1);

        M3Fwd_Demand := (PRG_01_Diagnostics.FB_Joystick_0.AxisCmdX.Direction = 1);
        M3Rev_Demand := (PRG_01_Diagnostics.FB_Joystick_0.AxisCmdX.Direction = -1);
    ELSE
        // 💡 Détection de mouvement en cours (pour verrouillage croisé)
        WinchMoving := M1Fwd_Demand OR M1Rev_Demand OR M2Fwd_Demand OR M2Rev_Demand OR CoupledFwd_Demand OR CoupledRev_Demand;

        // 🔒 Verrouillage d'aiguillage HMI : on ne démarre un mouvement que si aucun autre n'est en cours
        // 🔧 REX 2026-07-15 (2) : ex-tenue "AND SpeedRefPct > 0.1" retirée — rampe HMI locale
        // supprimée (M1/M2 pilotés via FB_Winch, PRG_06_WinchControl), qui gère désormais SEUL la
        // rampe et l'interlock de changement de sens (DirectionChangePending/DirectionChangeDelay,
        // voir FB_Winch.st) : plus besoin de tenir la demande le temps d'une décél locale ici.
        M1Fwd_Demand := GVL_IHM.IHM_MANU.M1_RelayFwd AND (NOT WinchMoving OR M1Fwd_Demand);
        M1Rev_Demand := GVL_IHM.IHM_MANU.M1_RelayRev AND (NOT WinchMoving OR M1Rev_Demand);
        M2Fwd_Demand := GVL_IHM.IHM_MANU.M2_RelayFwd AND (NOT WinchMoving OR M2Fwd_Demand);
        M2Rev_Demand := GVL_IHM.IHM_MANU.M2_RelayRev AND (NOT WinchMoving OR M2Rev_Demand);
        CoupledFwd_Demand := GVL_IHM.IHM_MANU.M1_M2_RelayFwd AND (NOT WinchMoving OR CoupledFwd_Demand);
        CoupledRev_Demand := GVL_IHM.IHM_MANU.M1_M2_RelayRev AND (NOT WinchMoving OR CoupledRev_Demand);

        M3Fwd_Demand := GVL_IHM.TranslationM3.ReqFwd;
        M3Rev_Demand := GVL_IHM.TranslationM3.ReqRev;
    END_IF;

    // 🔒 Sécurité démarrage : exige que toutes les commandes HMI et Joystick soient au repos (neutre) au démarrage
    IF NOT StartupNeutralOk THEN
        IF NOT GVL_IHM.IHM_MANU.M1_RelayFwd AND NOT GVL_IHM.IHM_MANU.M1_RelayRev
           AND NOT GVL_IHM.IHM_MANU.M2_RelayFwd AND NOT GVL_IHM.IHM_MANU.M2_RelayRev
           AND NOT GVL_IHM.IHM_MANU.M1_M2_RelayFwd AND NOT GVL_IHM.IHM_MANU.M1_M2_RelayRev
           AND NOT GVL_IHM.TranslationM3.ReqFwd AND NOT GVL_IHM.TranslationM3.ReqRev
           AND ABS(PRG_01_Diagnostics.FB_Joystick_0.AxisCmdX.SpeedRef) < 1.0
           AND ABS(PRG_01_Diagnostics.FB_Joystick_0.AxisCmdY.SpeedRef) < 1.0 THEN
            StartupNeutralOk := TRUE;
        END_IF;
    END_IF;

    IF NOT StartupNeutralOk THEN
        M1Fwd_Demand := FALSE;
        M1Rev_Demand := FALSE;
        M2Fwd_Demand := FALSE;
        M2Rev_Demand := FALSE;
        CoupledFwd_Demand := FALSE;
        CoupledRev_Demand := FALSE;
        M3Fwd_Demand := FALSE;
        M3Rev_Demand := FALSE;
    END_IF;

    // 🔧 REX 2026-07-15 (2) : ex-§5️⃣/§5bis/§6️⃣ (M1Fwd_Eff/M1Rev_Eff/M2Fwd_Eff/M2Rev_Eff/
    // SimM1Fwd_Eff.../décodage K1-K4 via instManuSpeedStep) RETIRÉS — M1/M2 pilotés désormais par
    // instWinchM1/instWinchM2 (PRG_06_WinchControl §1/§2/§6/§7), qui écrivent directement
    // PRG_10_Outputs.M1RelayFwd/M1RelayRev/M1SpeedContactor1-4/M1BrakeCmd (et M2) via §8 de ce
    // même fichier PRG_06 — AVANT que ce PRG_10_Outputs ne s'exécute (position 6 < 10). Plus besoin
    // de "Recopie vers les VAR_INPUT" ci-dessous pour M1/M2 (voir fin de fichier).

    // 🔧 REX 2026-07-16 : ex-§7️⃣ (M3Fwd_Eff/M3Rev_Eff, interlock local avec M3_StatusWord.7/.0 et
    // SafeStop) RETIRÉ — M3 piloté désormais par instTranslationM3 (PRG_07_TranslationControl
    // §1bis), qui gère nativement SafeStop (Enable réel désormais, voir PRG_03_Safety) et sa
    // propre state machine. Plus besoin d'interlock local ici (même principe que M1/M2, REX
    // 2026-07-15 (2) ci-dessus).

    // 8️⃣ Auxiliaires Hydrauliques (action maintenue IHM + interlock logique d'exclusion mutuelle)
    IF GVL_IHM.IHM_MANU.GridOpenCmd AND NOT GVL_IHM.IHM_MANU.GridCloseCmd AND PRG_00_Inputs.EmergencyStopOk THEN
        GridUp_RQ := TRUE;
        GridDown_RQ := FALSE;
    ELSIF GVL_IHM.IHM_MANU.GridCloseCmd AND NOT GVL_IHM.IHM_MANU.GridOpenCmd AND PRG_00_Inputs.EmergencyStopOk THEN
        GridUp_RQ := FALSE;
        GridDown_RQ := TRUE;
    ELSE
        GridUp_RQ := FALSE;
        GridDown_RQ := FALSE;
    END_IF;

    IF GVL_IHM.IHM_MANU.HelmetOpenCmd AND NOT GVL_IHM.IHM_MANU.HelmetCloseCmd AND PRG_00_Inputs.EmergencyStopOk THEN
        HelmetOpen_RQ := TRUE;
        HelmetClose_RQ := FALSE;
    ELSIF GVL_IHM.IHM_MANU.HelmetCloseCmd AND NOT GVL_IHM.IHM_MANU.HelmetOpenCmd AND PRG_00_Inputs.EmergencyStopOk THEN
        HelmetOpen_RQ := FALSE;
        HelmetClose_RQ := TRUE;
    ELSE
        HelmetOpen_RQ := FALSE;
        HelmetClose_RQ := FALSE;
    END_IF;

    // Démarrage automatique du groupe hydraulique si un mouvement auxiliaire est demandé et AU armé
    PRG_08_AuxiliaryControl.HydraulicPumpRunCmd := (GVL_IHM.IHM_MANU.GridOpenCmd
                                                 OR GVL_IHM.IHM_MANU.GridCloseCmd
                                                 OR GVL_IHM.IHM_MANU.HelmetOpenCmd
                                                 OR GVL_IHM.IHM_MANU.HelmetCloseCmd)
                                                 AND PRG_00_Inputs.EmergencyStopOk;

    // 🔧 REX 2026-07-15 (2) : plus de recopie M1/M2 ici — déjà écrites par PRG_06_WinchControl §8
    // (instWinchM1/instWinchM2.RelayFwd/RelayRev/Contactor1-4/BrakeCmd), AVANT ce PRG_10_Outputs
    // dans l'ordre de tâche (position 6 < 10), pour Auto ET Manu désormais.
    // 🔧 REX 2026-07-16 : idem pour TranslationBrakeCmd — plus de recopie ici, déjà écrite par
    // PRG_07_TranslationControl (instTranslationM3.BrakeCmd), AVANT ce PRG_10_Outputs (position
    // 7 < 10), pour Auto ET Manu désormais (voir fin de fichier).
ELSE
    // Nettoyage en cas de désactivation du mode Manu
    GridUp_RQ := FALSE;
    GridDown_RQ := FALSE;
    HelmetOpen_RQ := FALSE;
    HelmetClose_RQ := FALSE;
END_IF;

// ── Translation M3 — variateur EtherCAT AC600, mot de commande direct (PAS de relais) ──
// 🔧 REX 2026-07-16 : ex-bypass ManuActive (écriture directe M3_CommandWord=1/2) RETIRÉ — M3
// piloté désormais par instTranslationM3 (PRG_07_TranslationControl §1bis), pour Auto ET Manu,
// même principe que M1/M2 (PRG_06_WinchControl §8, REX 2026-07-15 (2)).
M3_CommandWord         := PRG_07_TranslationControl.instTranslationM3.DriveControlWord;
M3_SetpointFrequencyHz := REAL_TO_UINT(PRG_07_TranslationControl.instTranslationM3.DriveFreqRefHz * 100.0);
// 🔧 DriveActualFreqHz / DriveCommReady / DrivePowerReady : écrits une seule fois, en
// PRG_09_Supervision (GVL_IHM.TranslationM3), valables Auto ET Manu — ex-doublons IHM_MANU
// M3_FreqActual/M3_CommandWordMonitor/M3_StatusWordMonitor/M3_CommReady/M3_PowerReady retirés.

// Relais de direction M3 obsolètes forcés à FALSE
M3_RelayFwd_DQ := FALSE;
M3_RelayRev_DQ := FALSE;

// 9️⃣ Enregistrement de l'état précédent (pour le cycle suivant)
LastM1Fwd      := GVL_IHM.IHM_MANU.M1_RelayFwd;
LastM1Rev      := GVL_IHM.IHM_MANU.M1_RelayRev;
LastM2Fwd      := GVL_IHM.IHM_MANU.M2_RelayFwd;
LastM2Rev      := GVL_IHM.IHM_MANU.M2_RelayRev;
LastCoupledFwd := GVL_IHM.IHM_MANU.M1_M2_RelayFwd;
LastCoupledRev := GVL_IHM.IHM_MANU.M1_M2_RelayRev;
LastM3Fwd      := GVL_IHM.TranslationM3.ReqFwd;
LastM3Rev      := GVL_IHM.TranslationM3.ReqRev;
// ─────────  Fin modification IHM_MANU  ─────────

// 🪝 ─── WINCH M1 — lit les VAR_INPUT de PRG_10_Outputs, écrit les I/O réels ────
instM1RelayFwd(Command := M1RelayFwd);
M1_RelayFwd_DQ := instM1RelayFwd.State;

instM1RelayRev(Command := M1RelayRev);
M1_RelayRev_DQ := instM1RelayRev.State;

instM1SpeedContactor1(Command := M1SpeedContactor1);
M1_SpeedContactor_1_DQ := instM1SpeedContactor1.State;

instM1SpeedContactor2(Command := M1SpeedContactor2);
M1_SpeedContactor_2_DQ := instM1SpeedContactor2.State;

instM1SpeedContactor3(Command := M1SpeedContactor3);
M1_SpeedContactor_3_DQ := instM1SpeedContactor3.State;

instM1SpeedContactor4(Command := M1SpeedContactor4);
M1_SpeedContactor_4_DQ := instM1SpeedContactor4.State;

instM1BrakeCmd(Command := M1BrakeCmd);
M1_BrakeCmd_RQ := instM1BrakeCmd.State;

// 🪝 ─── WINCH M2 ──────────────────────────────────────────────────────────
instM2RelayFwd(Command := M2RelayFwd);
M2_RelayFwd_DQ := instM2RelayFwd.State;

instM2RelayRev(Command := M2RelayRev);
M2_RelayRev_DQ := instM2RelayRev.State;

instM2SpeedContactor1(Command := M2SpeedContactor1);
M2_SpeedContactor_1_DQ := instM2SpeedContactor1.State;

instM2SpeedContactor2(Command := M2SpeedContactor2);
M2_SpeedContactor_2_DQ := instM2SpeedContactor2.State;

instM2SpeedContactor3(Command := M2SpeedContactor3);
M2_SpeedContactor_3_DQ := instM2SpeedContactor3.State;

instM2SpeedContactor4(Command := M2SpeedContactor4);
M2_SpeedContactor_4_DQ := instM2SpeedContactor4.State;

instM2BrakeCmd(Command := M2BrakeCmd);
M2_BrakeCmd_RQ := instM2BrakeCmd.State;

// ↔️ ─── TRANSLATION M3 ────────────────────────────────────────────────────────
instTranslationBrakeCmd(Command := TranslationBrakeCmd);
M3_BrakeCmd_RQ := instTranslationBrakeCmd.State;

// ─── 🧨 COUPURE PUISSANCE AMONT REDONDANTE (Série physique, commande parallèle) ────────
// Calcul du besoin de coupure amont (intégrant le bypass en mode IHM_MANU)
PowerCutOffReq := (ManuActive AND PowerCutOffActive_Eff)
                  OR (NOT ManuActive AND (PRG_03_Safety.instSafetyWinchM1.PowerCutOff
                                       OR PRG_03_Safety.instSafetyWinchM2.PowerCutOff
                                       OR PRG_03_Safety.instSafetyTranslationM3.PowerCutOff));

// Appel du bloc Safety global pour la boucle d'urgence
instSafetyEmergencyManagement(
    Enable := TRUE,
    Reset := PRG_09_Supervision.FaultMachineReset_IHM,
    ArmRequest := GVL_IHM.Modes.CmdEmergencyArming,
    EmergencyChain := PRG_00_Inputs.EmergencyChain,
    EmergencyStopOk := PRG_00_Inputs.EmergencyStopOk,
    PowerCutOffRequest := PowerCutOffReq,
    CmdEmergencyCutOff := NOT ManuActive AND GVL_IHM.Modes.CmdEmergencyCutOff
);

// Affectation des sorties physiques et logiques de coupure/réarmement
PowerCutOff_A_RQ := instSafetyEmergencyManagement.PowerCutOff_A_RQ;
PowerCutOff_B_RQ := instSafetyEmergencyManagement.PowerCutOff_B_RQ;
EmergencyArming_RQ := instSafetyEmergencyManagement.EmergencyArming_RQ;

// Copie des états de diagnostic vers la supervision IHM
EmergencyArmingPulseActive   := instSafetyEmergencyManagement.EmergencyArming_RQ;
EmergencyArmingLockoutActive := instSafetyEmergencyManagement.EmergencyArmingLockoutActive;
ArmingSeqStep                := instSafetyEmergencyManagement.ArmingSeqStep;
RedundancyTestFailed         := instSafetyEmergencyManagement.RedundancyTestFailed;
EmergencyArmingFailed        := instSafetyEmergencyManagement.EmergencyArmingFailed;

(* ---- PRG_IP.st ---- *)
(* ═══════════════════════════════════════════════════════════════
   💻 PRG_IP — Configuration / Diagnostic Ethernet / IP
   ───────────────────────────────────────────────────────────────
   Note : Programme exécuté en tâche de fond ou asynchrone.
   Le bloc de configuration de l'IP est actuellement stubbé / commenté.
   ═══════════════════════════════════════════════════════════════ *)
PROGRAM PRG_IP
VAR
    // SetNetworkConfig_0 : SetNetworkConfig; (* Configuration IP commentée par défaut *)
END_VAR

// Pas d'implémentation active (toutes les configurations sont figées ou gérées par l'OS automate).
